# EPICS autosave request: 1.5.0/debian-12/7.0.10/modules/ADCore-ee039d2/db/NDCircularBuff_settings.req
$(P)$(R)TriggerA
$(P)$(R)TriggerB
$(P)$(R)TriggerCalc
$(P)$(R)PreCount
$(P)$(R)PostCount
$(P)$(R)PresetTriggerCount
$(P)$(R)FlushOnSoftTrg
file "NDPluginBase_settings.req", P=$(P), R=$(R)
